(* IEC 61131-3 sources: tsplc/examples/bottling-line/raw-st/src/publication, 2 files *)

(* ---- GVL_Example.st ---- *)
{attribute 'qualified_only'}
VAR_GLOBAL CONSTANT
	Description : STRING := 'Bottling line raw ST example';
END_VAR

(* ---- PRG_Publish.declaration.st ---- *)
PROGRAM PRG_Publish
VAR
	Heartbeat : UDINT;
END_VAR
